(* Logix 5000 project; controller R400_500_XLS vendor 1 type 14 code 216 rev 31.11; software revision 31.01; part 30 of 32 *)
(* tags used below, declared in another part *)
   Alarm : SINT;   // Wait 3 seconds
   CalibData : UDT_SCALE[8];
   Chem_Pump : UDT_CHEM_PUMP[4];   // Chemical Pump flow rate
   FC45_NextMaintDate : DINT[3];   // Next maintenance due date
   FINAL_RINSE_MAX_NBR : INT;   // Maximum nimber of final rinse
   M : DINT[5];   // Memory Bits
   MaxPressRecord : REAL;
   NeutralizantPump : SINT;
   OneShot : DINT[1];
   print_Footer_template : STRING[7];   // Template for the cycle footer
   print_Header_template : STRING[6];   // Template for the cycle header
   PrintCalibdata : STRING[9];
   printNeutralization : STRING[5];
   PrintSensorName : STRING[7];
   printTreatString : STRING[85];   // Treatment String
   rIn_WSH61 : REAL;
   sCRLF : STRING;
   sOut_WSH61 : STRING;
   sPrntArray : STRING[300];   // Printer String Array
   SRE3_Serial_Number : STRING;   // Serial number
   String_Temp : STRING;
   Tmr : TIMER[107];
   WSH41_Total_time : STRING;
   WSH61_Footer : STRING[6];   // The footer being transferred to the print queue.
   CalibCounter : SINT;
   Cfg_11_Modules : BOOL;
   ChemicalName : STRING[9];   // Used by HMI
   CR2Mode : SINT;   // 0= Cycle complete dry contact 1= External pure water valve
   CycleCounter : DINT;
   DateTime : DINT[7];
   ENABLE : BOOL;   // Enable bit
   FC45_NbCycBeforeMaint : DINT;
   iDelayBeforeFillingAuthAlarmMM : DINT;
   iDelayBeforeFillingAuthAlarmSS : DINT;
   iInactivityLogoutTime : DINT;   // Inactivity Logout Time In Minutes
   iPWClosingDelayMM : DINT;
   iPWClosingDelaySS : DINT;
   iSCADACycleCompleteTimeHr : INT;
   iSCADACycleCompleteTimeMin : INT;
   iSCADACycleCompleteTimeSec : INT;
   Language_English : STRING;
   Non_Vented_with_Dry_Option : BOOL;
   NonVented_Without_Dry_Option : BOOL;
   NumInput : UDT_NUMERIC_INPUT[65];   // Numeric input
   NumInputReal : UDT_NUMERIC_INPUT_REAL[17];
   PressureUnit : BOOL;   // Pressure Unit 0=PSIG 1=BAR
   PrintHardware : STRING[29];
   PrintIndex : DINT;
   PrintSystemOption : STRING[29];
   sChangeLanguage : STRING;   // jplv09
   sCycleCounter : STRING;
   SPV_19 : BOOL;   // Screen 80 Enabled/Disabled Pump pressure monitoring
   sTime : STRING;   // String current time
   Tpb : DINT[11];
   Unit : Hrdwre;   // Unit Configuration
   UnLoad : Doors;
   Vented_with_Dry_Option : BOOL;
(* MainProgram, continued *)

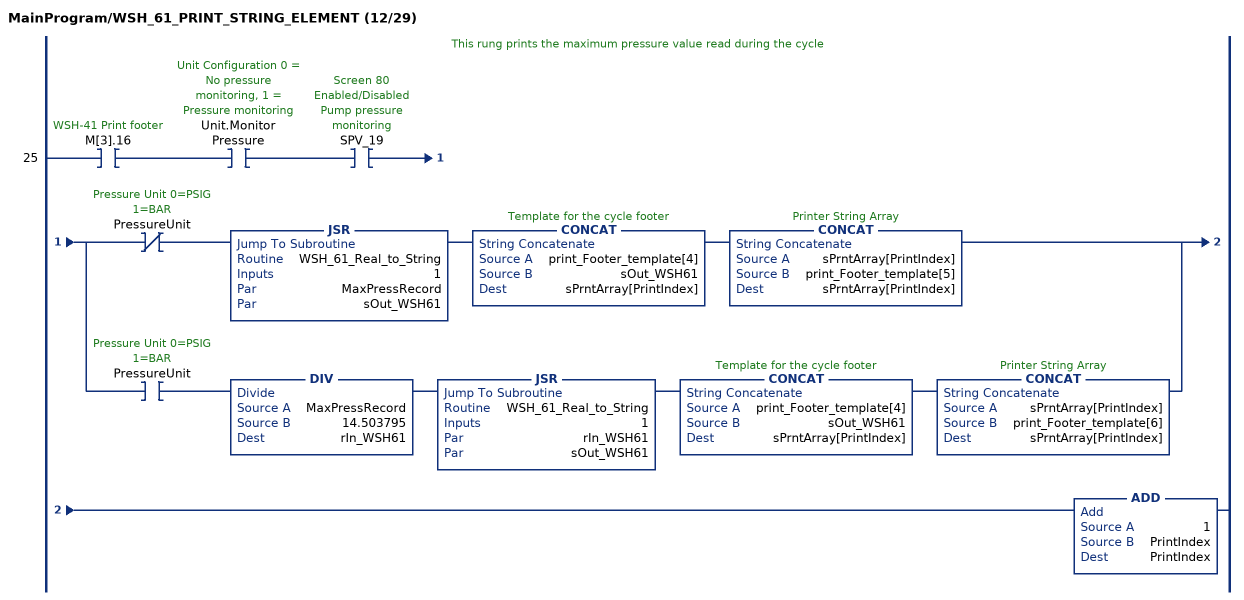
   [picture p617: MainProgram/WSH_61_PRINT_STRING_ELEMENT rungs 25-25]
   // This rung prints the maximum pressure value read during the cycle
   25: XIC(M[3].16)XIC(Unit.MonitorPressure)XIC(SPV_19)[XIO(PressureUnit) JSR(WSH_61_Real_to_String,1,MaxPressRecord,sOut_WSH61) CONCAT(print_Footer_template[4],sOut_WSH61,sPrntArray[PrintIndex]) CONCAT(sPrntArray[PrintIndex],print_Footer_template[5],sPrntArray[PrintIndex]) ,XIC(PressureUnit) DIV(MaxPressRecord,14.503795,rIn_WSH61) JSR(WSH_61_Real_to_String,1,rIn_WSH61,sOut_WSH61) CONCAT(print_Footer_template[4],sOut_WSH61,sPrntArray[PrintIndex]) CONCAT(sPrntArray[PrintIndex],print_Footer_template[6],sPrntArray[PrintIndex]) ]ADD(1,PrintIndex,PrintIndex);
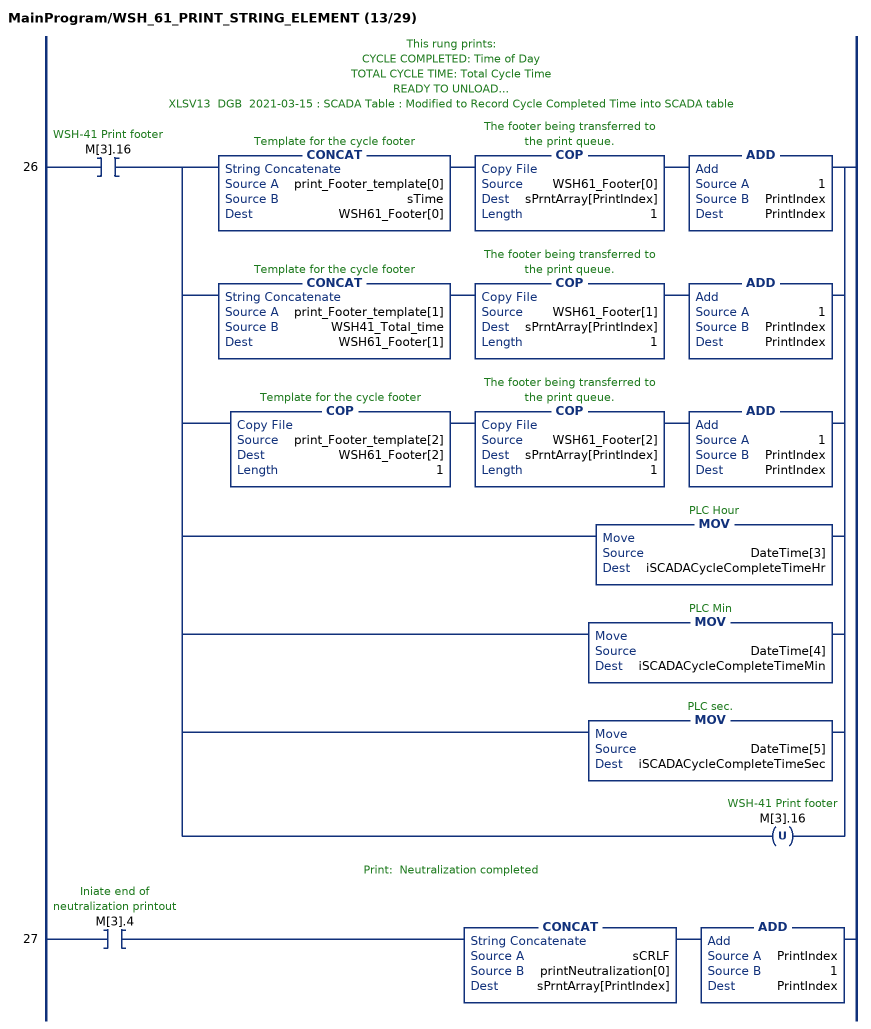
   // This rung prints:
   // CYCLE COMPLETED: Time of Day
   // TOTAL CYCLE TIME: Total Cycle Time
   // READY TO UNLOAD...
   // XLSV13  DGB  2021-03-15 : SCADA Table : Modified to Record Cycle Completed Time into SCADA table
   26: XIC(M[3].16)[CONCAT(print_Footer_template[0],sTime,WSH61_Footer[0]) COP(WSH61_Footer[0],sPrntArray[PrintIndex],1) ADD(1,PrintIndex,PrintIndex) ,CONCAT(print_Footer_template[1],WSH41_Total_time,WSH61_Footer[1]) COP(WSH61_Footer[1],sPrntArray[PrintIndex],1) ADD(1,PrintIndex,PrintIndex) ,COP(print_Footer_template[2],WSH61_Footer[2],1) COP(WSH61_Footer[2],sPrntArray[PrintIndex],1) ADD(1,PrintIndex,PrintIndex) ,[MOV(DateTime[3],iSCADACycleCompleteTimeHr) ,MOV(DateTime[4],iSCADACycleCompleteTimeMin) ,MOV(DateTime[5],iSCADACycleCompleteTimeSec) ] ,OTU(M[3].16) ];
   // Print:  Neutralization completed
   27: XIC(M[3].4)CONCAT(sCRLF,printNeutralization[0],sPrntArray[PrintIndex])ADD(PrintIndex,1,PrintIndex);
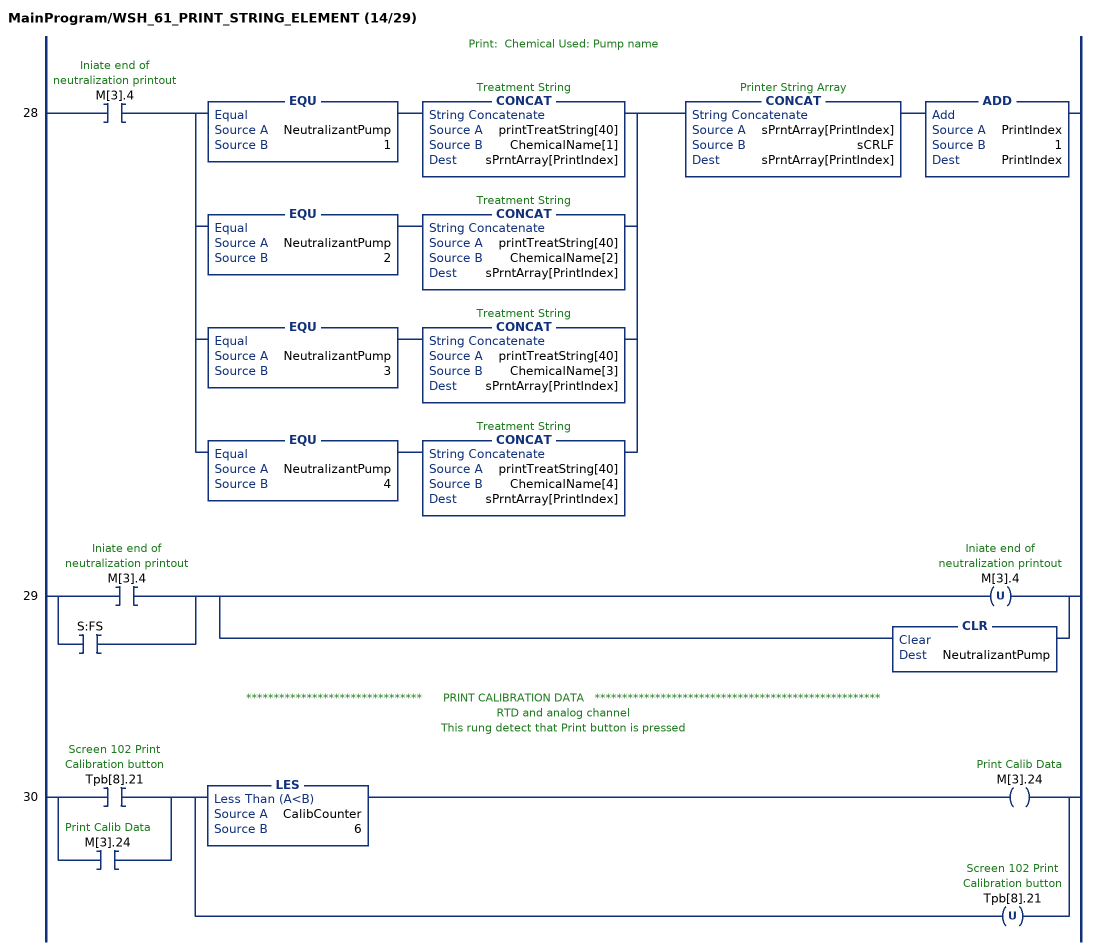
   // Print:  Chemical Used: Pump name
   28: XIC(M[3].4)[EQU(NeutralizantPump,1) CONCAT(printTreatString[40],ChemicalName[1],sPrntArray[PrintIndex]) ,EQU(NeutralizantPump,2) CONCAT(printTreatString[40],ChemicalName[2],sPrntArray[PrintIndex]) ,EQU(NeutralizantPump,3) CONCAT(printTreatString[40],ChemicalName[3],sPrntArray[PrintIndex]) ,EQU(NeutralizantPump,4) CONCAT(printTreatString[40],ChemicalName[4],sPrntArray[PrintIndex]) ]CONCAT(sPrntArray[PrintIndex],sCRLF,sPrntArray[PrintIndex])ADD(PrintIndex,1,PrintIndex);
   29: [XIC(M[3].4) ,XIC(S:FS) ][OTU(M[3].4) ,CLR(NeutralizantPump) ];
   // ********************************      PRINT CALIBRATION DATA   ****************************************************
   // RTD and analog channel
   // This rung detect that Print button is pressed
   30: [XIC(Tpb[8].21) ,XIC(M[3].24) ][LES(CalibCounter,6) OTE(M[3].24) ,OTU(Tpb[8].21) ];
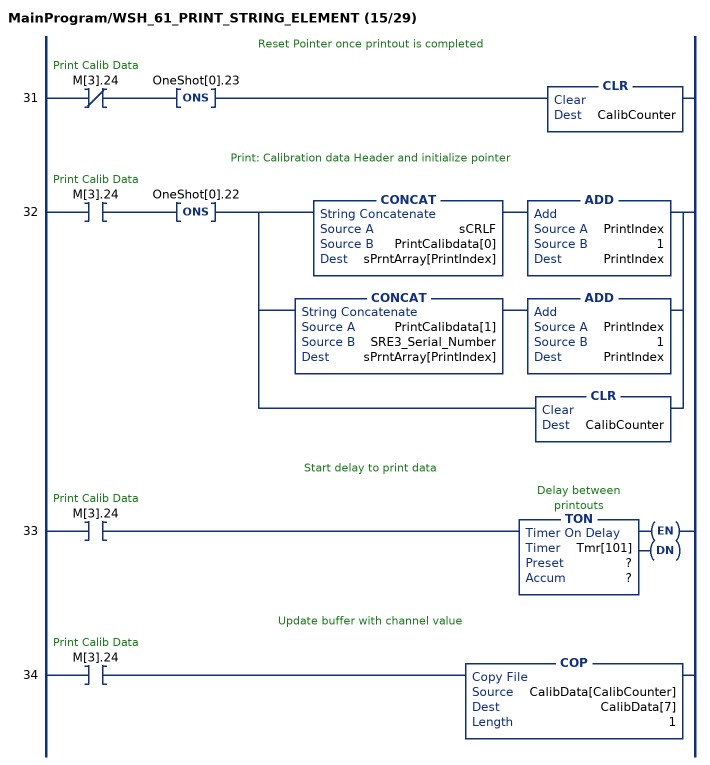
   // Reset Pointer once printout is completed
   31: XIO(M[3].24)ONS(OneShot[0].23)CLR(CalibCounter);
   // Print: Calibration data Header and initialize pointer
   32: XIC(M[3].24)ONS(OneShot[0].22)[CONCAT(sCRLF,PrintCalibdata[0],sPrntArray[PrintIndex]) ADD(PrintIndex,1,PrintIndex) ,CONCAT(PrintCalibdata[1],SRE3_Serial_Number,sPrntArray[PrintIndex]) ADD(PrintIndex,1,PrintIndex) ,CLR(CalibCounter) ];
   // Start delay to print data
   33: XIC(M[3].24)TON(Tmr[101],?,?);
   // Update buffer with channel value
   34: XIC(M[3].24)COP(CalibData[CalibCounter],CalibData[7],1);
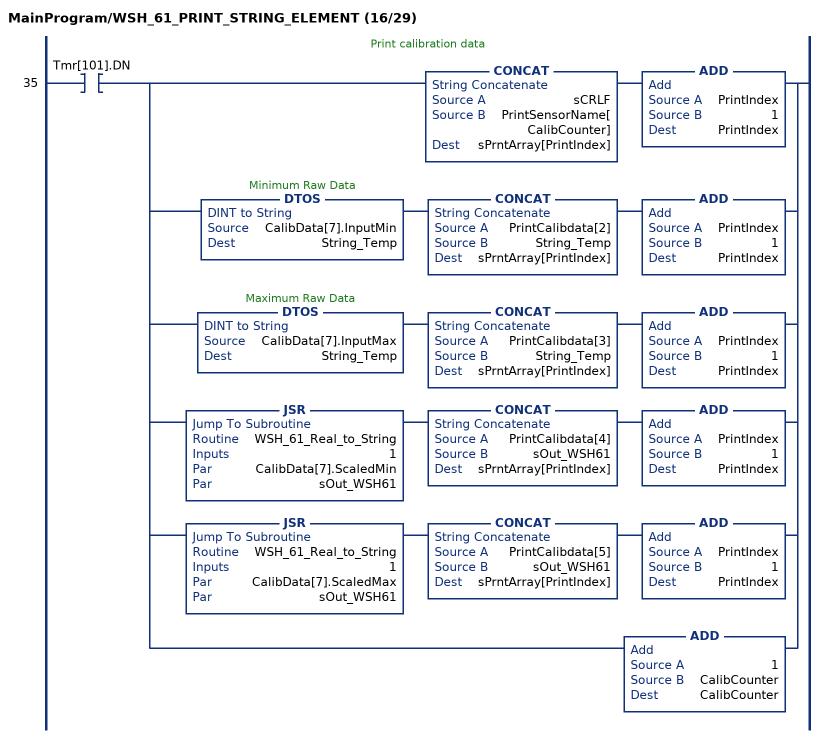
   // Print calibration data
   35: XIC(Tmr[101].DN)[CONCAT(sCRLF,PrintSensorName[CalibCounter],sPrntArray[PrintIndex]) ADD(PrintIndex,1,PrintIndex) ,DTOS(CalibData[7].InputMin,String_Temp) CONCAT(PrintCalibdata[2],String_Temp,sPrntArray[PrintIndex]) ADD(PrintIndex,1,PrintIndex) ,DTOS(CalibData[7].InputMax,String_Temp) CONCAT(PrintCalibdata[3],String_Temp,sPrntArray[PrintIndex]) ADD(PrintIndex,1,PrintIndex) ,JSR(WSH_61_Real_to_String,1,CalibData[7].ScaledMin,sOut_WSH61) CONCAT(PrintCalibdata[4],sOut_WSH61,sPrntArray[PrintIndex]) ADD(PrintIndex,1,PrintIndex) ,JSR(WSH_61_Real_to_String,1,CalibData[7].ScaledMax,sOut_WSH61) CONCAT(PrintCalibdata[5],sOut_WSH61,sPrntArray[PrintIndex]) ADD(PrintIndex,1,PrintIndex) ,ADD(1,CalibCounter,CalibCounter) ];
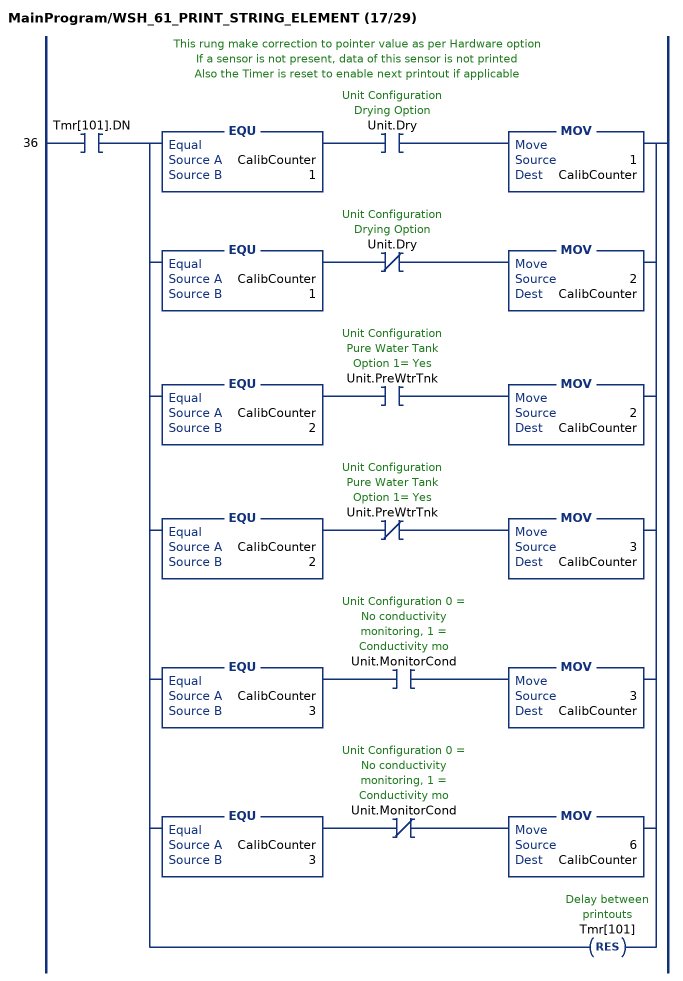
   // This rung make correction to pointer value as per Hardware option
   // If a sensor is not present, data of this sensor is not printed
   // Also the Timer is reset to enable next printout if applicable
   36: XIC(Tmr[101].DN)[EQU(CalibCounter,1) XIC(Unit.Dry) MOV(1,CalibCounter) ,EQU(CalibCounter,1) XIO(Unit.Dry) MOV(2,CalibCounter) ,EQU(CalibCounter,2) XIC(Unit.PreWtrTnk) MOV(2,CalibCounter) ,EQU(CalibCounter,2) XIO(Unit.PreWtrTnk) MOV(3,CalibCounter) ,EQU(CalibCounter,3) XIC(Unit.MonitorCond) MOV(3,CalibCounter) ,EQU(CalibCounter,3) XIO(Unit.MonitorCond) MOV(6,CalibCounter) ,RES(Tmr[101]) ];
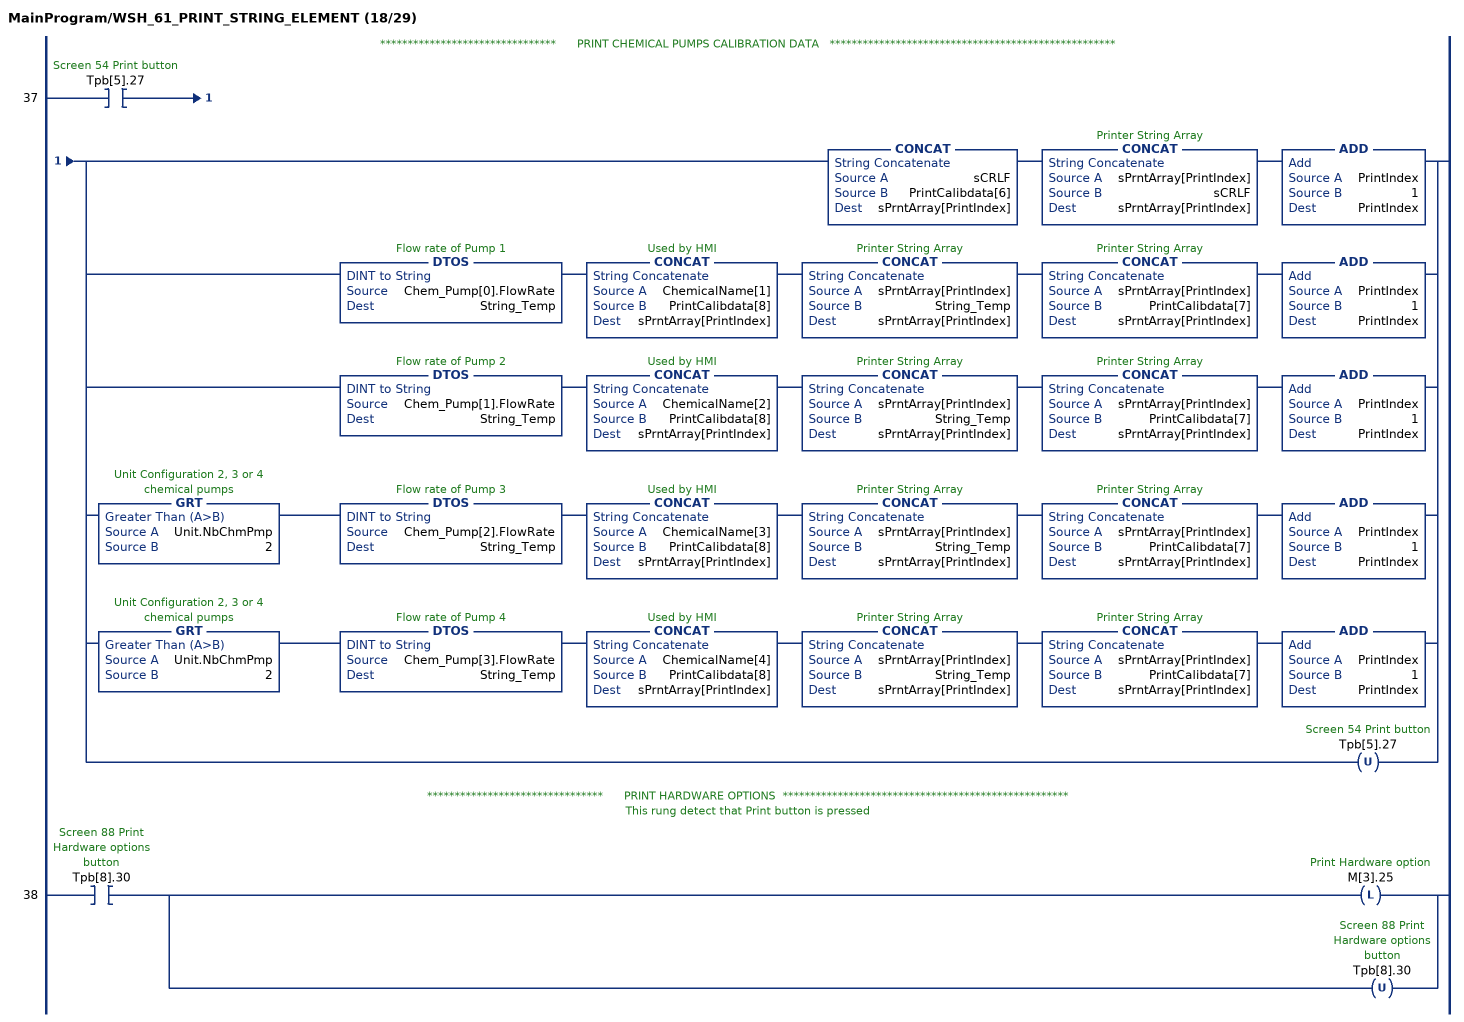
   // ********************************      PRINT CHEMICAL PUMPS CALIBRATION DATA   ****************************************************
   37: XIC(Tpb[5].27)[CONCAT(sCRLF,PrintCalibdata[6],sPrntArray[PrintIndex]) CONCAT(sPrntArray[PrintIndex],sCRLF,sPrntArray[PrintIndex]) ADD(PrintIndex,1,PrintIndex) ,DTOS(Chem_Pump[0].FlowRate,String_Temp) CONCAT(ChemicalName[1],PrintCalibdata[8],sPrntArray[PrintIndex]) CONCAT(sPrntArray[PrintIndex],String_Temp,sPrntArray[PrintIndex]) CONCAT(sPrntArray[PrintIndex],PrintCalibdata[7],sPrntArray[PrintIndex]) ADD(PrintIndex,1,PrintIndex) ,DTOS(Chem_Pump[1].FlowRate,String_Temp) CONCAT(ChemicalName[2],PrintCalibdata[8],sPrntArray[PrintIndex]) CONCAT(sPrntArray[PrintIndex],String_Temp,sPrntArray[PrintIndex]) CONCAT(sPrntArray[PrintIndex],PrintCalibdata[7],sPrntArray[PrintIndex]) ADD(PrintIndex,1,PrintIndex) ,GRT(Unit.NbChmPmp,2) DTOS(Chem_Pump[2].FlowRate,String_Temp) CONCAT(ChemicalName[3],PrintCalibdata[8],sPrntArray[PrintIndex]) CONCAT(sPrntArray[PrintIndex],String_Temp,sPrntArray[PrintIndex]) CONCAT(sPrntArray[PrintIndex],PrintCalibdata[7],sPrntArray[PrintIndex]) ADD(PrintIndex,1,PrintIndex) ,GRT(Unit.NbChmPmp,2) DTOS(Chem_Pump[3].FlowRate,String_Temp) CONCAT(ChemicalName[4],PrintCalibdata[8],sPrntArray[PrintIndex]) CONCAT(sPrntArray[PrintIndex],String_Temp,sPrntArray[PrintIndex]) CONCAT(sPrntArray[PrintIndex],PrintCalibdata[7],sPrntArray[PrintIndex]) ADD(PrintIndex,1,PrintIndex) ,OTU(Tpb[5].27) ];
   // ********************************      PRINT HARDWARE OPTIONS  ****************************************************
   // This rung detect that Print button is pressed
   38: XIC(Tpb[8].30)[OTL(M[3].25) ,OTU(Tpb[8].30) ];
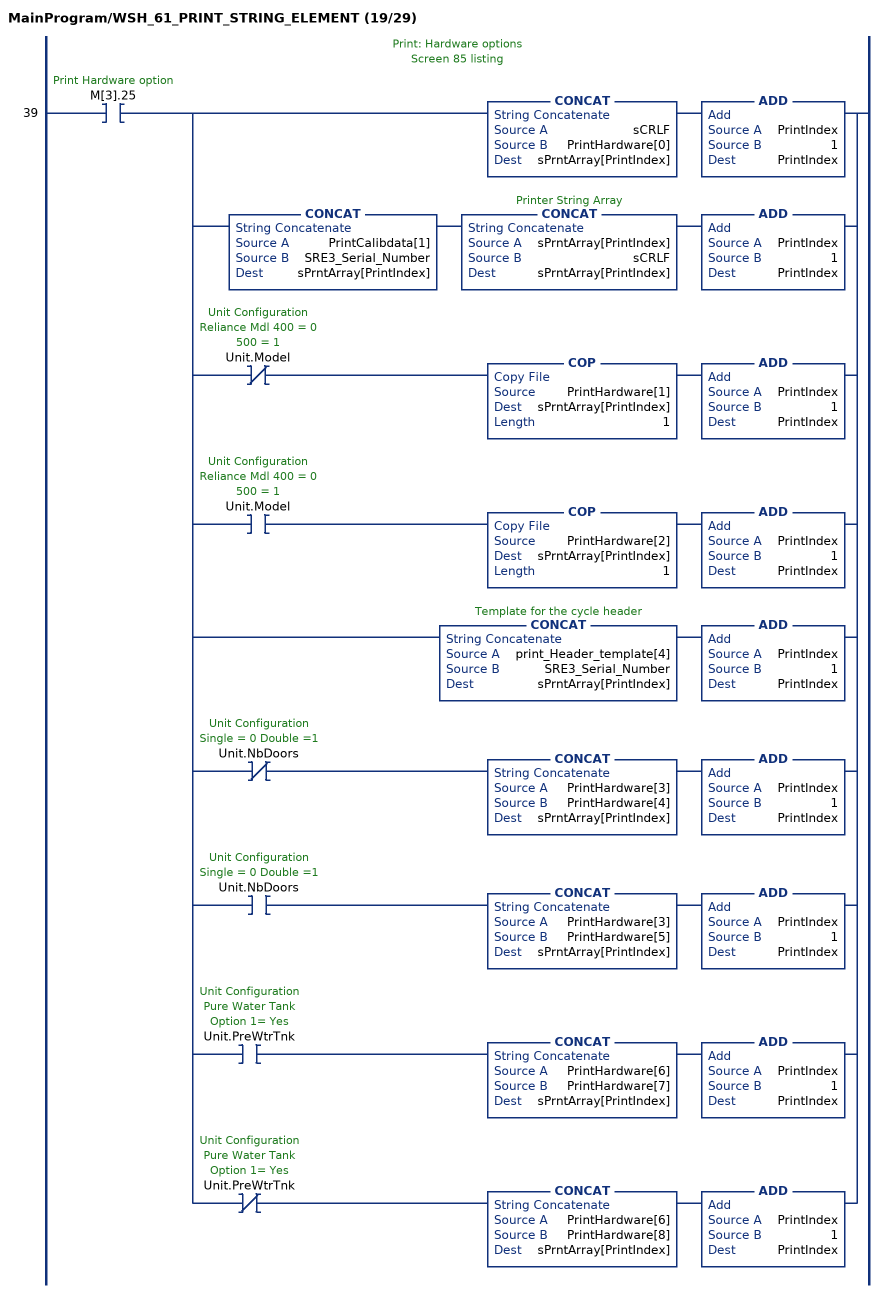
   // Print: Hardware options
   // Screen 85 listing
   39: XIC(M[3].25)[CONCAT(sCRLF,PrintHardware[0],sPrntArray[PrintIndex]) ADD(PrintIndex,1,PrintIndex) ,CONCAT(PrintCalibdata[1],SRE3_Serial_Number,sPrntArray[PrintIndex]) CONCAT(sPrntArray[PrintIndex],sCRLF,sPrntArray[PrintIndex]) ADD(PrintIndex,1,PrintIndex) ,XIO(Unit.Model) COP(PrintHardware[1],sPrntArray[PrintIndex],1) ADD(PrintIndex,1,PrintIndex) ,XIC(Unit.Model) COP(PrintHardware[2],sPrntArray[PrintIndex],1) ADD(PrintIndex,1,PrintIndex) ,CONCAT(print_Header_template[4],SRE3_Serial_Number,sPrntArray[PrintIndex]) ADD(PrintIndex,1,PrintIndex) ,XIO(Unit.NbDoors) CONCAT(PrintHardware[3],PrintHardware[4],sPrntArray[PrintIndex]) ADD(PrintIndex,1,PrintIndex) ,XIC(Unit.NbDoors) CONCAT(PrintHardware[3],PrintHardware[5],sPrntArray[PrintIndex]) ADD(PrintIndex,1,PrintIndex) ,XIC(Unit.PreWtrTnk) CONCAT(PrintHardware[6],PrintHardware[7],sPrntArray[PrintIndex]) ADD(PrintIndex,1,PrintIndex) ,XIO(Unit.PreWtrTnk) CONCAT(PrintHardware[6],PrintHardware[8],sPrntArray[PrintIndex]) ADD(PrintIndex,1,PrintIndex) ];
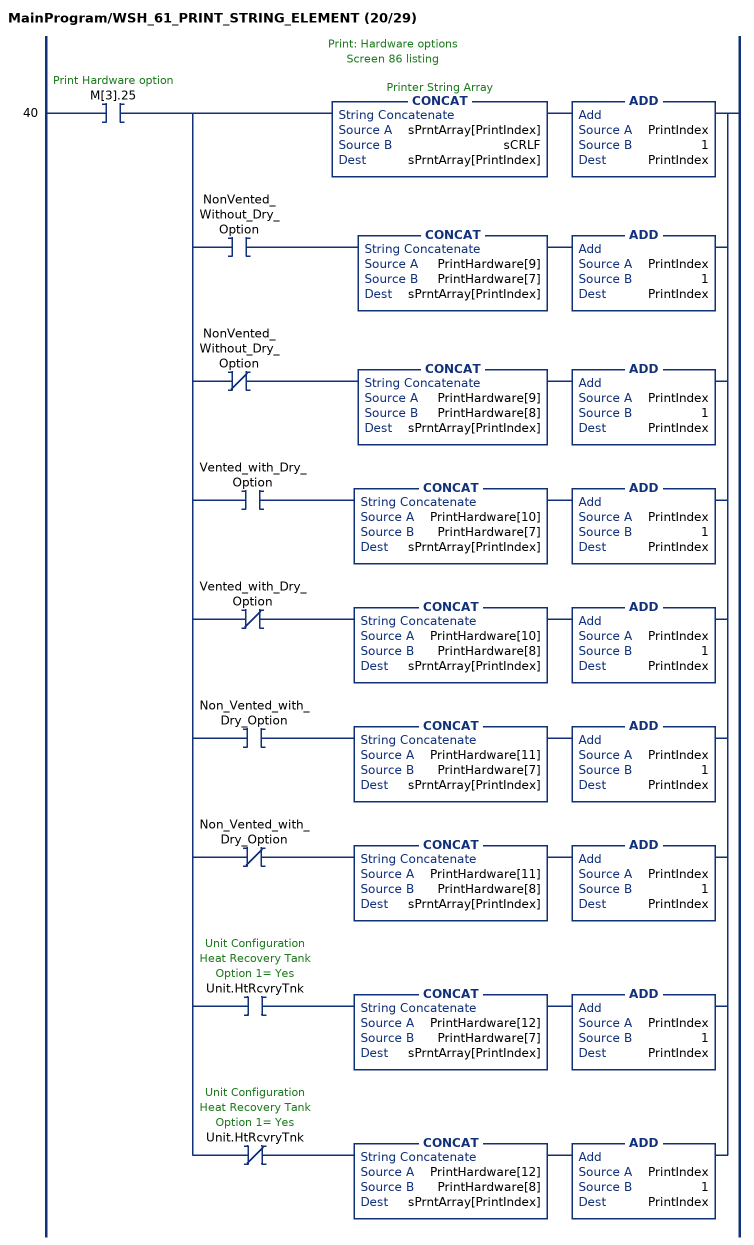
   // Print: Hardware options
   // Screen 86 listing
   40: XIC(M[3].25)[CONCAT(sPrntArray[PrintIndex],sCRLF,sPrntArray[PrintIndex]) ADD(PrintIndex,1,PrintIndex) ,XIC(NonVented_Without_Dry_Option) CONCAT(PrintHardware[9],PrintHardware[7],sPrntArray[PrintIndex]) ADD(PrintIndex,1,PrintIndex) ,XIO(NonVented_Without_Dry_Option) CONCAT(PrintHardware[9],PrintHardware[8],sPrntArray[PrintIndex]) ADD(PrintIndex,1,PrintIndex) ,XIC(Vented_with_Dry_Option) CONCAT(PrintHardware[10],PrintHardware[7],sPrntArray[PrintIndex]) ADD(PrintIndex,1,PrintIndex) ,XIO(Vented_with_Dry_Option) CONCAT(PrintHardware[10],PrintHardware[8],sPrntArray[PrintIndex]) ADD(PrintIndex,1,PrintIndex) ,XIC(Non_Vented_with_Dry_Option) CONCAT(PrintHardware[11],PrintHardware[7],sPrntArray[PrintIndex]) ADD(PrintIndex,1,PrintIndex) ,XIO(Non_Vented_with_Dry_Option) CONCAT(PrintHardware[11],PrintHardware[8],sPrntArray[PrintIndex]) ADD(PrintIndex,1,PrintIndex) ,XIC(Unit.HtRcvryTnk) CONCAT(PrintHardware[12],PrintHardware[7],sPrntArray[PrintIndex]) ADD(PrintIndex,1,PrintIndex) ,XIO(Unit.HtRcvryTnk) CONCAT(PrintHardware[12],PrintHardware[8],sPrntArray[PrintIndex]) ADD(PrintIndex,1,PrintIndex) ];
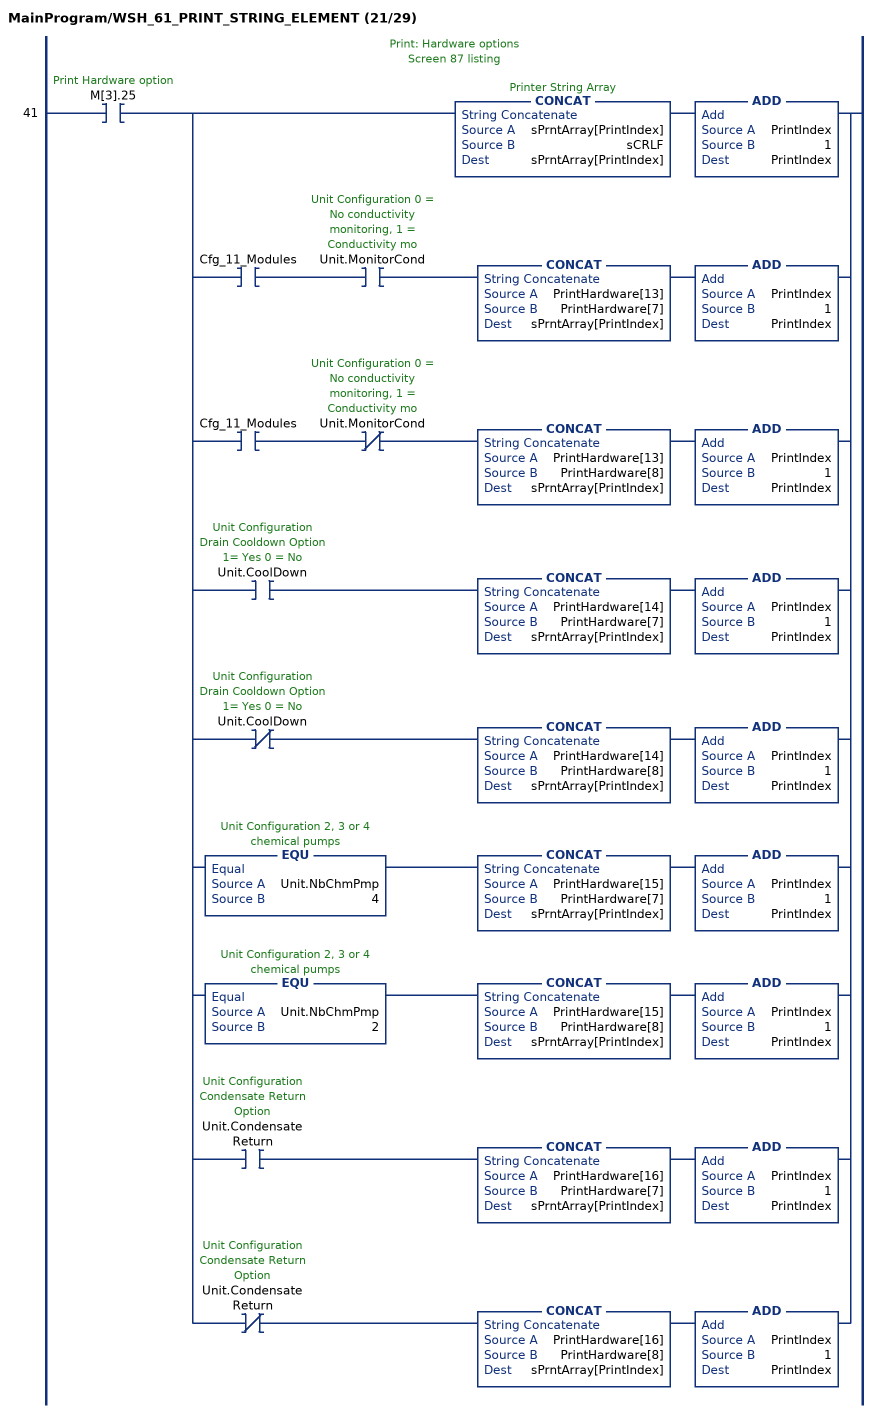
   // Print: Hardware options
   // Screen 87 listing
   41: XIC(M[3].25)[CONCAT(sPrntArray[PrintIndex],sCRLF,sPrntArray[PrintIndex]) ADD(PrintIndex,1,PrintIndex) ,XIC(Cfg_11_Modules) XIC(Unit.MonitorCond) CONCAT(PrintHardware[13],PrintHardware[7],sPrntArray[PrintIndex]) ADD(PrintIndex,1,PrintIndex) ,XIC(Cfg_11_Modules) XIO(Unit.MonitorCond) CONCAT(PrintHardware[13],PrintHardware[8],sPrntArray[PrintIndex]) ADD(PrintIndex,1,PrintIndex) ,XIC(Unit.CoolDown) CONCAT(PrintHardware[14],PrintHardware[7],sPrntArray[PrintIndex]) ADD(PrintIndex,1,PrintIndex) ,XIO(Unit.CoolDown) CONCAT(PrintHardware[14],PrintHardware[8],sPrntArray[PrintIndex]) ADD(PrintIndex,1,PrintIndex) ,EQU(Unit.NbChmPmp,4) CONCAT(PrintHardware[15],PrintHardware[7],sPrntArray[PrintIndex]) ADD(PrintIndex,1,PrintIndex) ,EQU(Unit.NbChmPmp,2) CONCAT(PrintHardware[15],PrintHardware[8],sPrntArray[PrintIndex]) ADD(PrintIndex,1,PrintIndex) ,XIC(Unit.CondensateReturn) CONCAT(PrintHardware[16],PrintHardware[7],sPrntArray[PrintIndex]) ADD(PrintIndex,1,PrintIndex) ,XIO(Unit.CondensateReturn) CONCAT(PrintHardware[16],PrintHardware[8],sPrntArray[PrintIndex]) ADD(PrintIndex,1,PrintIndex) ];
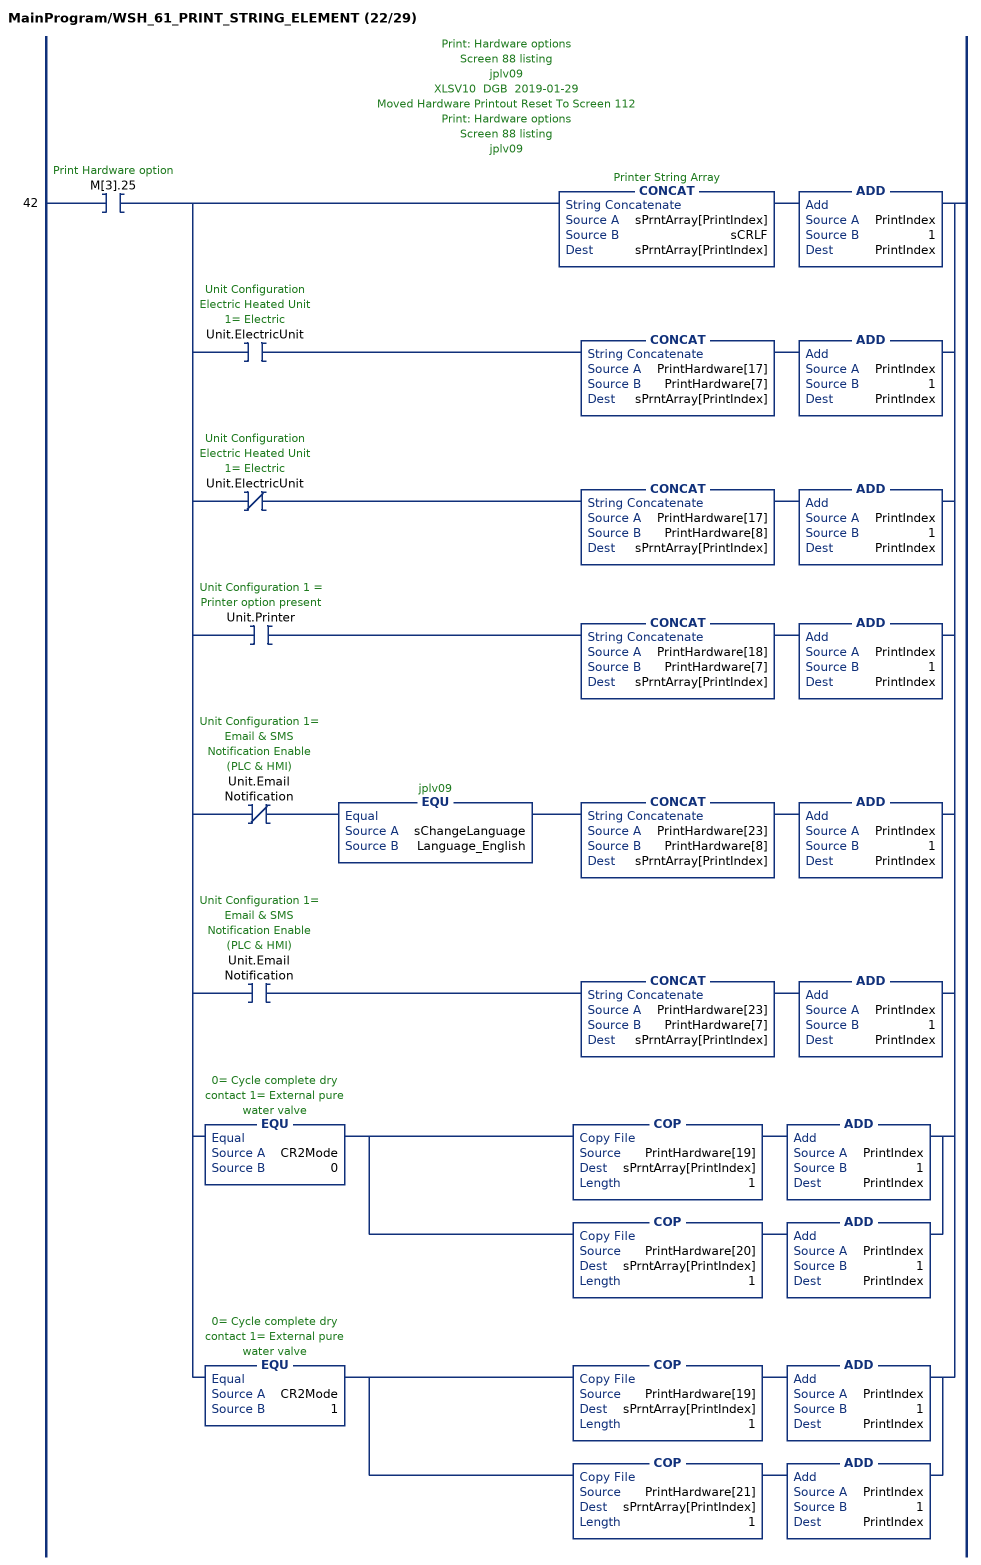
   // Print: Hardware options
   // Screen 88 listing
   // jplv09
   // XLSV10  DGB  2019-01-29
   // Moved Hardware Printout Reset To Screen 112
   // Print: Hardware options
   // Screen 88 listing
   // jplv09
   42: XIC(M[3].25)[CONCAT(sPrntArray[PrintIndex],sCRLF,sPrntArray[PrintIndex]) ADD(PrintIndex,1,PrintIndex) ,XIC(Unit.ElectricUnit) CONCAT(PrintHardware[17],PrintHardware[7],sPrntArray[PrintIndex]) ADD(PrintIndex,1,PrintIndex) ,XIO(Unit.ElectricUnit) CONCAT(PrintHardware[17],PrintHardware[8],sPrntArray[PrintIndex]) ADD(PrintIndex,1,PrintIndex) ,XIC(Unit.Printer) CONCAT(PrintHardware[18],PrintHardware[7],sPrntArray[PrintIndex]) ADD(PrintIndex,1,PrintIndex) ,XIO(Unit.EmailNotification) EQU(sChangeLanguage,Language_English) CONCAT(PrintHardware[23],PrintHardware[8],sPrntArray[PrintIndex]) ADD(PrintIndex,1,PrintIndex) ,XIC(Unit.EmailNotification) CONCAT(PrintHardware[23],PrintHardware[7],sPrntArray[PrintIndex]) ADD(PrintIndex,1,PrintIndex) ,EQU(CR2Mode,0) [COP(PrintHardware[19],sPrntArray[PrintIndex],1) ADD(PrintIndex,1,PrintIndex) ,COP(PrintHardware[20],sPrntArray[PrintIndex],1) ADD(PrintIndex,1,PrintIndex) ] ,EQU(CR2Mode,1) [COP(PrintHardware[19],sPrntArray[PrintIndex],1) ADD(PrintIndex,1,PrintIndex) ,COP(PrintHardware[21],sPrntArray[PrintIndex],1) ADD(PrintIndex,1,PrintIndex) ] ];
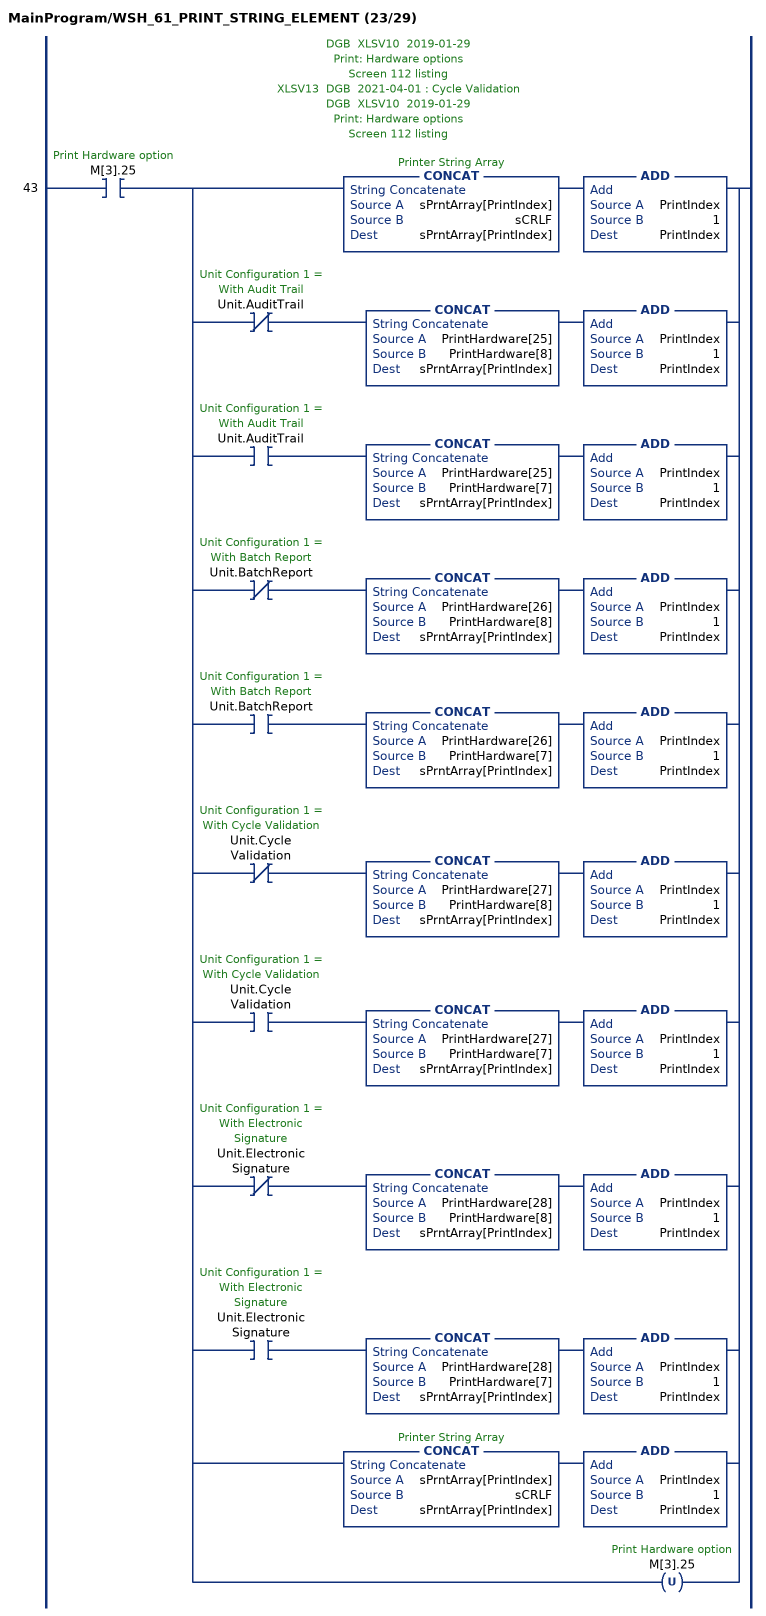
   // DGB  XLSV10  2019-01-29
   // Print: Hardware options
   // Screen 112 listing
   // XLSV13  DGB  2021-04-01 : Cycle Validation
   // DGB  XLSV10  2019-01-29
   // Print: Hardware options
   // Screen 112 listing
   43: XIC(M[3].25)[CONCAT(sPrntArray[PrintIndex],sCRLF,sPrntArray[PrintIndex]) ADD(PrintIndex,1,PrintIndex) ,XIO(Unit.AuditTrail) CONCAT(PrintHardware[25],PrintHardware[8],sPrntArray[PrintIndex]) ADD(PrintIndex,1,PrintIndex) ,XIC(Unit.AuditTrail) CONCAT(PrintHardware[25],PrintHardware[7],sPrntArray[PrintIndex]) ADD(PrintIndex,1,PrintIndex) ,XIO(Unit.BatchReport) CONCAT(PrintHardware[26],PrintHardware[8],sPrntArray[PrintIndex]) ADD(PrintIndex,1,PrintIndex) ,XIC(Unit.BatchReport) CONCAT(PrintHardware[26],PrintHardware[7],sPrntArray[PrintIndex]) ADD(PrintIndex,1,PrintIndex) ,XIO(Unit.CycleValidation) CONCAT(PrintHardware[27],PrintHardware[8],sPrntArray[PrintIndex]) ADD(PrintIndex,1,PrintIndex) ,XIC(Unit.CycleValidation) CONCAT(PrintHardware[27],PrintHardware[7],sPrntArray[PrintIndex]) ADD(PrintIndex,1,PrintIndex) ,XIO(Unit.ElectronicSignature) CONCAT(PrintHardware[28],PrintHardware[8],sPrntArray[PrintIndex]) ADD(PrintIndex,1,PrintIndex) ,XIC(Unit.ElectronicSignature) CONCAT(PrintHardware[28],PrintHardware[7],sPrntArray[PrintIndex]) ADD(PrintIndex,1,PrintIndex) ,CONCAT(sPrntArray[PrintIndex],sCRLF,sPrntArray[PrintIndex]) ADD(PrintIndex,1,PrintIndex) ,OTU(M[3].25) ];
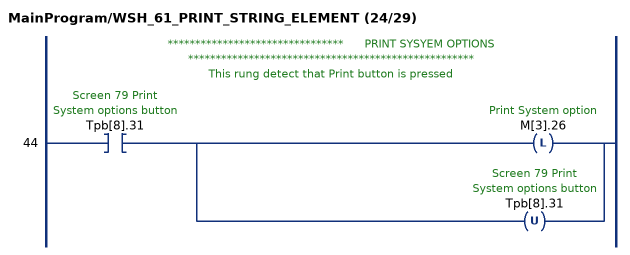
   // ********************************      PRINT SYSYEM OPTIONS  ****************************************************
   // This rung detect that Print button is pressed
   44: XIC(Tpb[8].31)[OTL(M[3].26) ,OTU(Tpb[8].31) ];
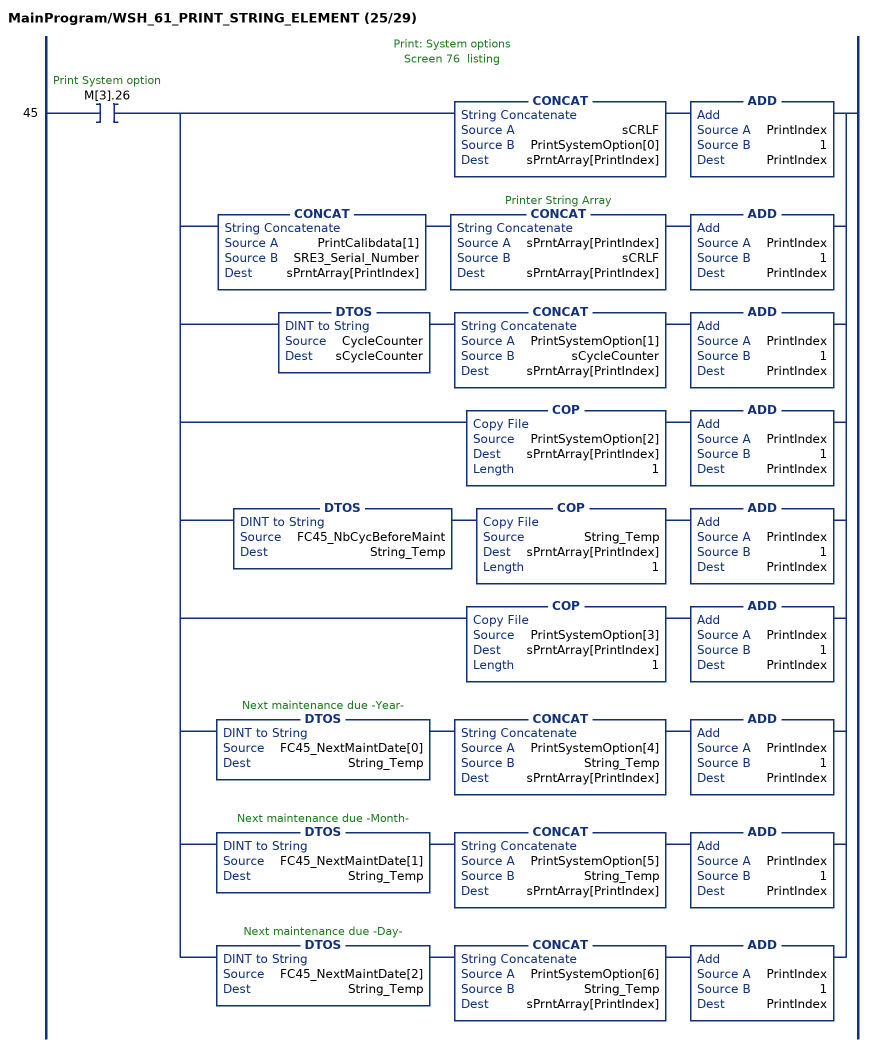
   // Print: System options
   // Screen 76  listing
   45: XIC(M[3].26)[CONCAT(sCRLF,PrintSystemOption[0],sPrntArray[PrintIndex]) ADD(PrintIndex,1,PrintIndex) ,CONCAT(PrintCalibdata[1],SRE3_Serial_Number,sPrntArray[PrintIndex]) CONCAT(sPrntArray[PrintIndex],sCRLF,sPrntArray[PrintIndex]) ADD(PrintIndex,1,PrintIndex) ,DTOS(CycleCounter,sCycleCounter) CONCAT(PrintSystemOption[1],sCycleCounter,sPrntArray[PrintIndex]) ADD(PrintIndex,1,PrintIndex) ,COP(PrintSystemOption[2],sPrntArray[PrintIndex],1) ADD(PrintIndex,1,PrintIndex) ,DTOS(FC45_NbCycBeforeMaint,String_Temp) COP(String_Temp,sPrntArray[PrintIndex],1) ADD(PrintIndex,1,PrintIndex) ,COP(PrintSystemOption[3],sPrntArray[PrintIndex],1) ADD(PrintIndex,1,PrintIndex) ,DTOS(FC45_NextMaintDate[0],String_Temp) CONCAT(PrintSystemOption[4],String_Temp,sPrntArray[PrintIndex]) ADD(PrintIndex,1,PrintIndex) ,DTOS(FC45_NextMaintDate[1],String_Temp) CONCAT(PrintSystemOption[5],String_Temp,sPrntArray[PrintIndex]) ADD(PrintIndex,1,PrintIndex) ,DTOS(FC45_NextMaintDate[2],String_Temp) CONCAT(PrintSystemOption[6],String_Temp,sPrntArray[PrintIndex]) ADD(PrintIndex,1,PrintIndex) ];
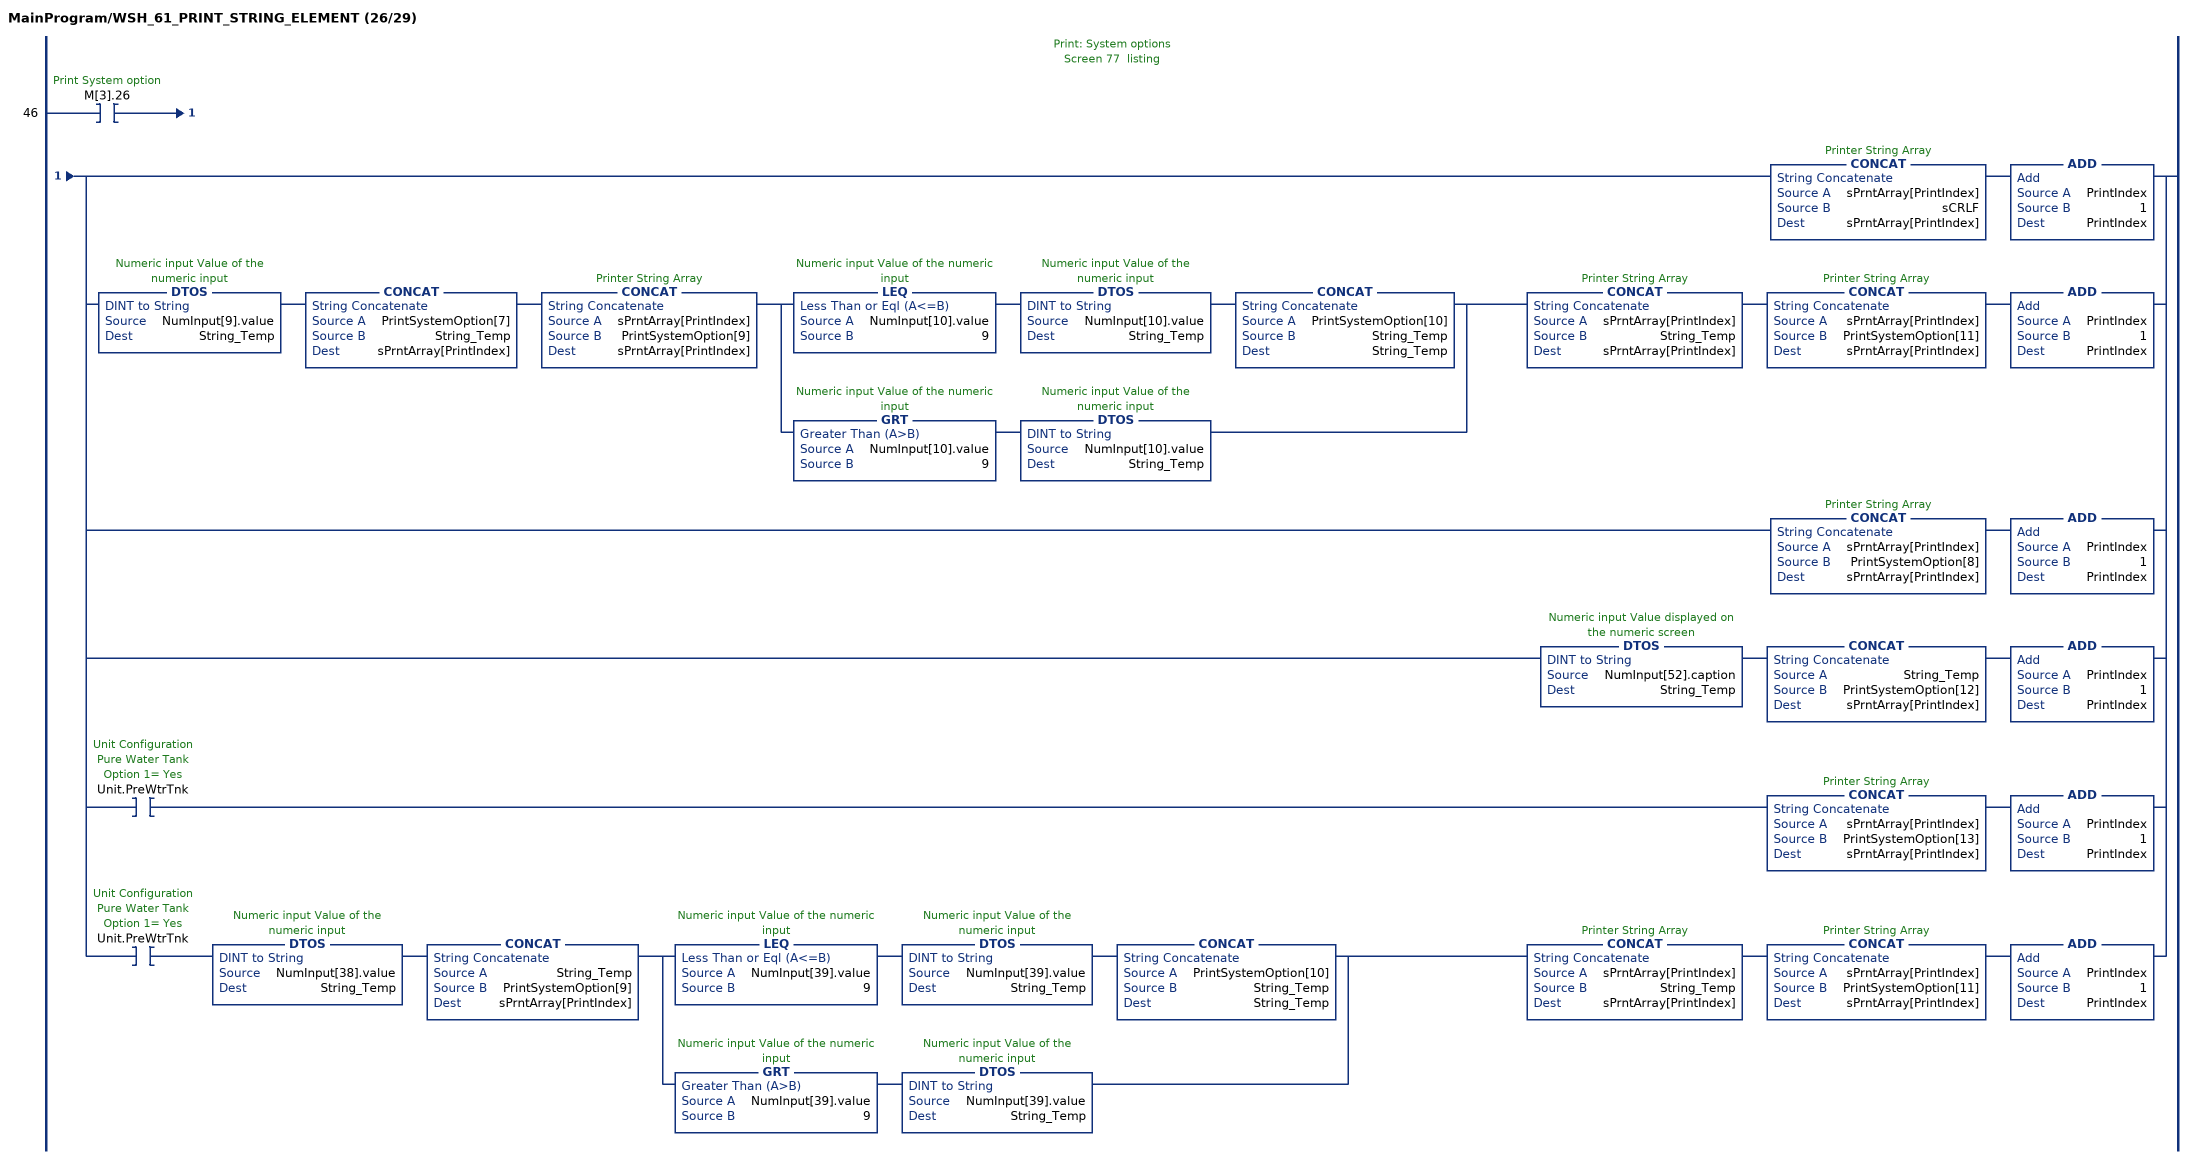
   // Print: System options
   // Screen 77  listing
   46: XIC(M[3].26)[CONCAT(sPrntArray[PrintIndex],sCRLF,sPrntArray[PrintIndex]) ADD(PrintIndex,1,PrintIndex) ,DTOS(NumInput[9].value,String_Temp) CONCAT(PrintSystemOption[7],String_Temp,sPrntArray[PrintIndex]) CONCAT(sPrntArray[PrintIndex],PrintSystemOption[9],sPrntArray[PrintIndex]) [LEQ(NumInput[10].value,9) DTOS(NumInput[10].value,String_Temp) CONCAT(PrintSystemOption[10],String_Temp,String_Temp) ,GRT(NumInput[10].value,9) DTOS(NumInput[10].value,String_Temp) ] CONCAT(sPrntArray[PrintIndex],String_Temp,sPrntArray[PrintIndex]) CONCAT(sPrntArray[PrintIndex],PrintSystemOption[11],sPrntArray[PrintIndex]) ADD(PrintIndex,1,PrintIndex) ,CONCAT(sPrntArray[PrintIndex],PrintSystemOption[8],sPrntArray[PrintIndex]) ADD(PrintIndex,1,PrintIndex) ,DTOS(NumInput[52].caption,String_Temp) CONCAT(String_Temp,PrintSystemOption[12],sPrntArray[PrintIndex]) ADD(PrintIndex,1,PrintIndex) ,XIC(Unit.PreWtrTnk) CONCAT(sPrntArray[PrintIndex],PrintSystemOption[13],sPrntArray[PrintIndex]) ADD(PrintIndex,1,PrintIndex) ,XIC(Unit.PreWtrTnk) DTOS(NumInput[38].value,String_Temp) CONCAT(String_Temp,PrintSystemOption[9],sPrntArray[PrintIndex]) [LEQ(NumInput[39].value,9) DTOS(NumInput[39].value,String_Temp) CONCAT(PrintSystemOption[10],String_Temp,String_Temp) ,GRT(NumInput[39].value,9) DTOS(NumInput[39].value,String_Temp) ] CONCAT(sPrntArray[PrintIndex],String_Temp,sPrntArray[PrintIndex]) CONCAT(sPrntArray[PrintIndex],PrintSystemOption[11],sPrntArray[PrintIndex]) ADD(PrintIndex,1,PrintIndex) ];
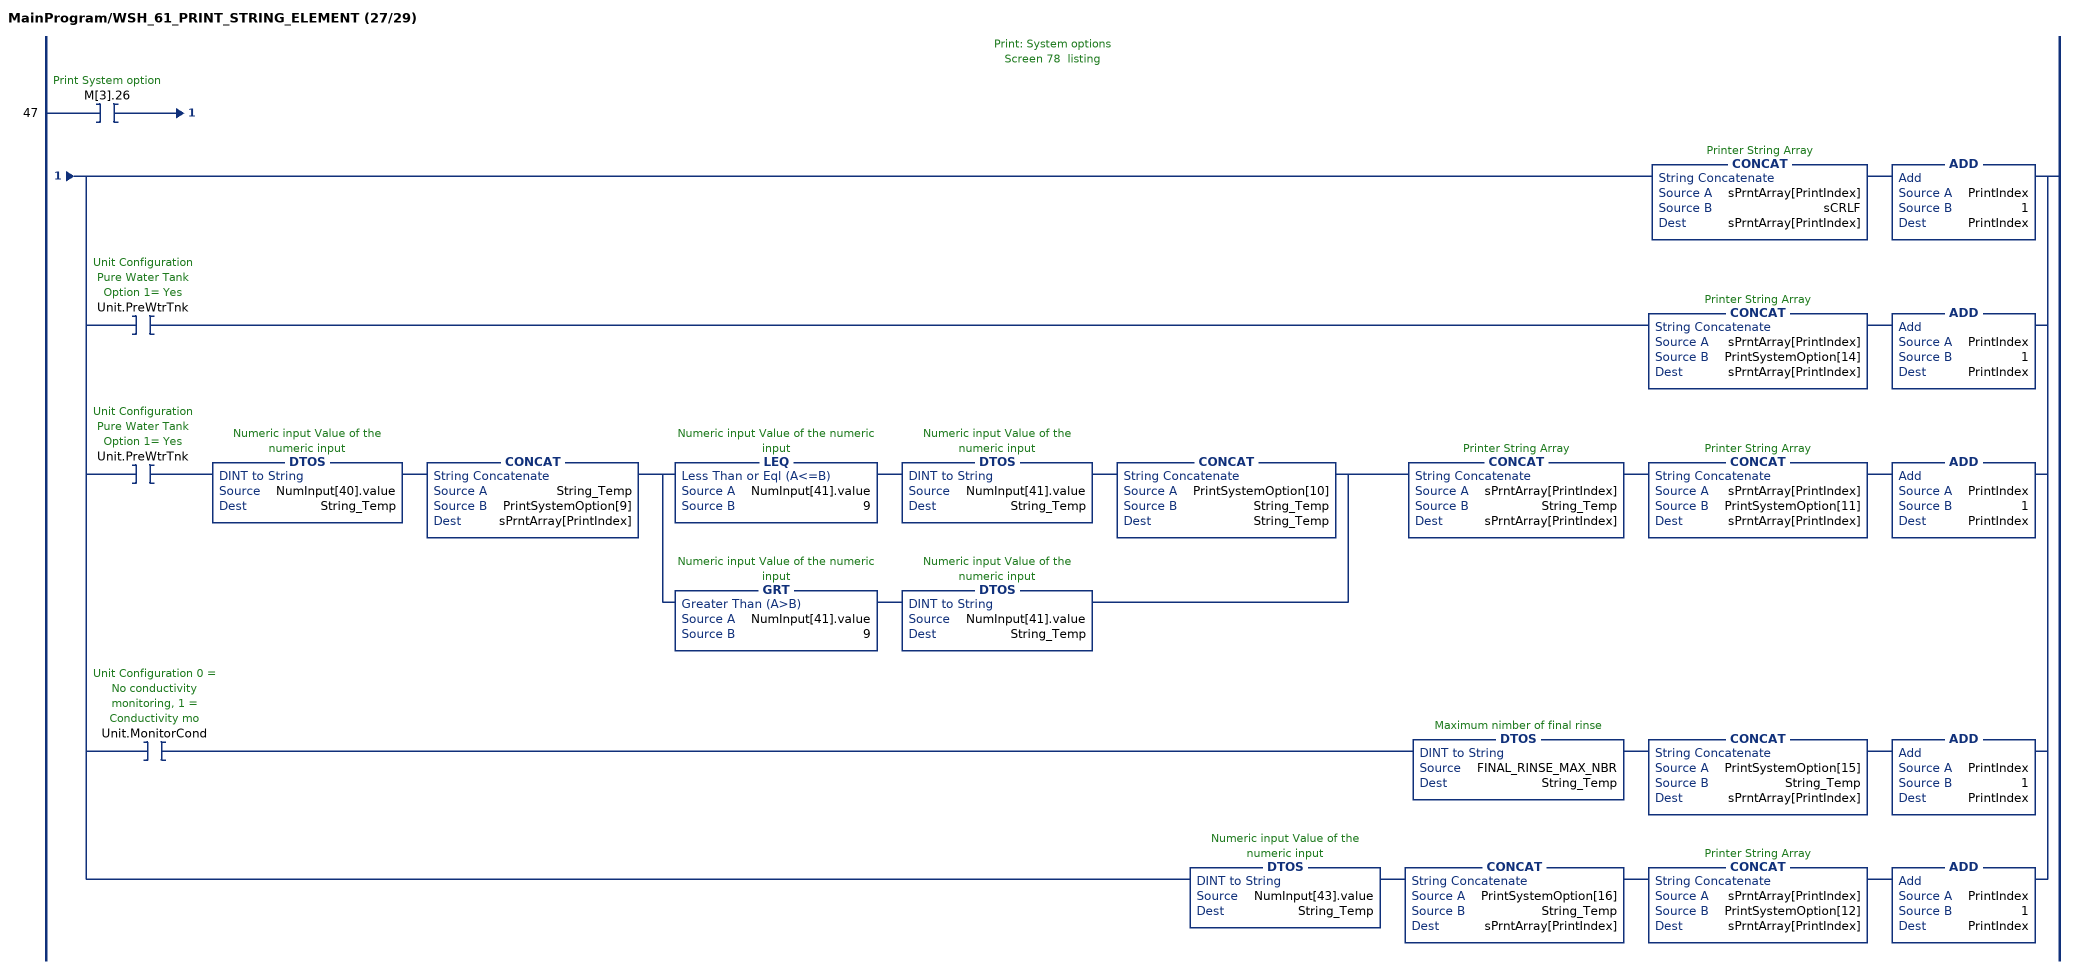
   // Print: System options
   // Screen 78  listing
   47: XIC(M[3].26)[CONCAT(sPrntArray[PrintIndex],sCRLF,sPrntArray[PrintIndex]) ADD(PrintIndex,1,PrintIndex) ,XIC(Unit.PreWtrTnk) CONCAT(sPrntArray[PrintIndex],PrintSystemOption[14],sPrntArray[PrintIndex]) ADD(PrintIndex,1,PrintIndex) ,XIC(Unit.PreWtrTnk) DTOS(NumInput[40].value,String_Temp) CONCAT(String_Temp,PrintSystemOption[9],sPrntArray[PrintIndex]) [LEQ(NumInput[41].value,9) DTOS(NumInput[41].value,String_Temp) CONCAT(PrintSystemOption[10],String_Temp,String_Temp) ,GRT(NumInput[41].value,9) DTOS(NumInput[41].value,String_Temp) ] CONCAT(sPrntArray[PrintIndex],String_Temp,sPrntArray[PrintIndex]) CONCAT(sPrntArray[PrintIndex],PrintSystemOption[11],sPrntArray[PrintIndex]) ADD(PrintIndex,1,PrintIndex) ,XIC(Unit.MonitorCond) DTOS(FINAL_RINSE_MAX_NBR,String_Temp) CONCAT(PrintSystemOption[15],String_Temp,sPrntArray[PrintIndex]) ADD(PrintIndex,1,PrintIndex) ,DTOS(NumInput[43].value,String_Temp) CONCAT(PrintSystemOption[16],String_Temp,sPrntArray[PrintIndex]) CONCAT(sPrntArray[PrintIndex],PrintSystemOption[12],sPrntArray[PrintIndex]) ADD(PrintIndex,1,PrintIndex) ];
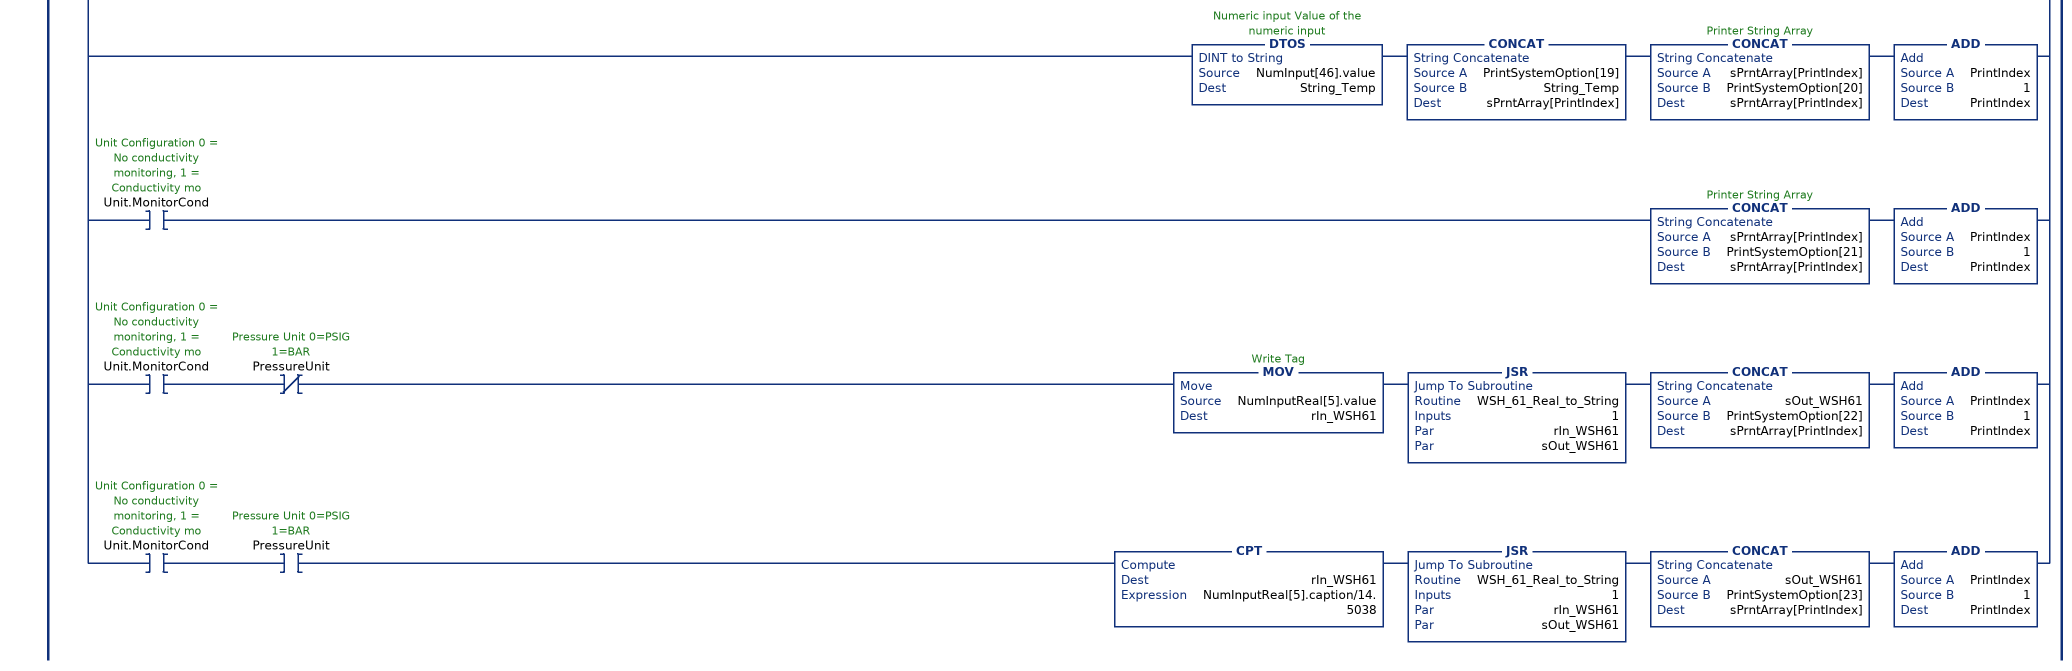
   // Print: System options
   // Screen 79  listing
   // XLSV10  DGB  2019-01-29
   // Moved End of System Option Printout in Screen 114
   48: XIC(M[3].26)[CONCAT(sPrntArray[PrintIndex],sCRLF,sPrntArray[PrintIndex]) ADD(PrintIndex,1,PrintIndex) ,CONCAT(sPrntArray[PrintIndex],PrintSystemOption[17],sPrntArray[PrintIndex]) ADD(PrintIndex,1,PrintIndex) ,DTOS(NumInput[44].value,String_Temp) CONCAT(String_Temp,PrintSystemOption[9],sPrntArray[PrintIndex]) [LEQ(NumInput[45].value,9) DTOS(NumInput[45].value,String_Temp) CONCAT(PrintSystemOption[10],String_Temp,String_Temp) ,GRT(NumInput[45].value,9) DTOS(NumInput[45].value,String_Temp) ] CONCAT(sPrntArray[PrintIndex],String_Temp,sPrntArray[PrintIndex]) CONCAT(sPrntArray[PrintIndex],PrintSystemOption[11],sPrntArray[PrintIndex]) ADD(PrintIndex,1,PrintIndex) ,XIC(Unit.Dry) CONCAT(sPrntArray[PrintIndex],PrintSystemOption[18],sPrntArray[PrintIndex]) ADD(PrintIndex,1,PrintIndex) ,XIC(Unit.Dry) DTOS(NumInput[47].value,String_Temp) CONCAT(String_Temp,PrintSystemOption[9],sPrntArray[PrintIndex]) [LEQ(NumInput[48].value,9) DTOS(NumInput[48].value,String_Temp) CONCAT(PrintSystemOption[10],String_Temp,String_Temp) ,GRT(NumInput[48].value,9) DTOS(NumInput[48].value,String_Temp) ] CONCAT(sPrntArray[PrintIndex],String_Temp,sPrntArray[PrintIndex]) CONCAT(sPrntArray[PrintIndex],PrintSystemOption[11],sPrntArray[PrintIndex]) ADD(PrintIndex,1,PrintIndex) ,DTOS(NumInput[46].value,String_Temp) CONCAT(PrintSystemOption[19],String_Temp,sPrntArray[PrintIndex]) CONCAT(sPrntArray[PrintIndex],PrintSystemOption[20],sPrntArray[PrintIndex]) ADD(PrintIndex,1,PrintIndex) ,XIC(Unit.MonitorCond) CONCAT(sPrntArray[PrintIndex],PrintSystemOption[21],sPrntArray[PrintIndex]) ADD(PrintIndex,1,PrintIndex) ,XIC(Unit.MonitorCond) XIO(PressureUnit) MOV(NumInputReal[5].value,rIn_WSH61) JSR(WSH_61_Real_to_String,1,rIn_WSH61,sOut_WSH61) CONCAT(sOut_WSH61,PrintSystemOption[22],sPrntArray[PrintIndex]) ADD(PrintIndex,1,PrintIndex) ,XIC(Unit.MonitorCond) XIC(PressureUnit) CPT(rIn_WSH61,NumInputReal[5].caption/14.5038) JSR(WSH_61_Real_to_String,1,rIn_WSH61,sOut_WSH61) CONCAT(sOut_WSH61,PrintSystemOption[23],sPrntArray[PrintIndex]) ADD(PrintIndex,1,PrintIndex) ];
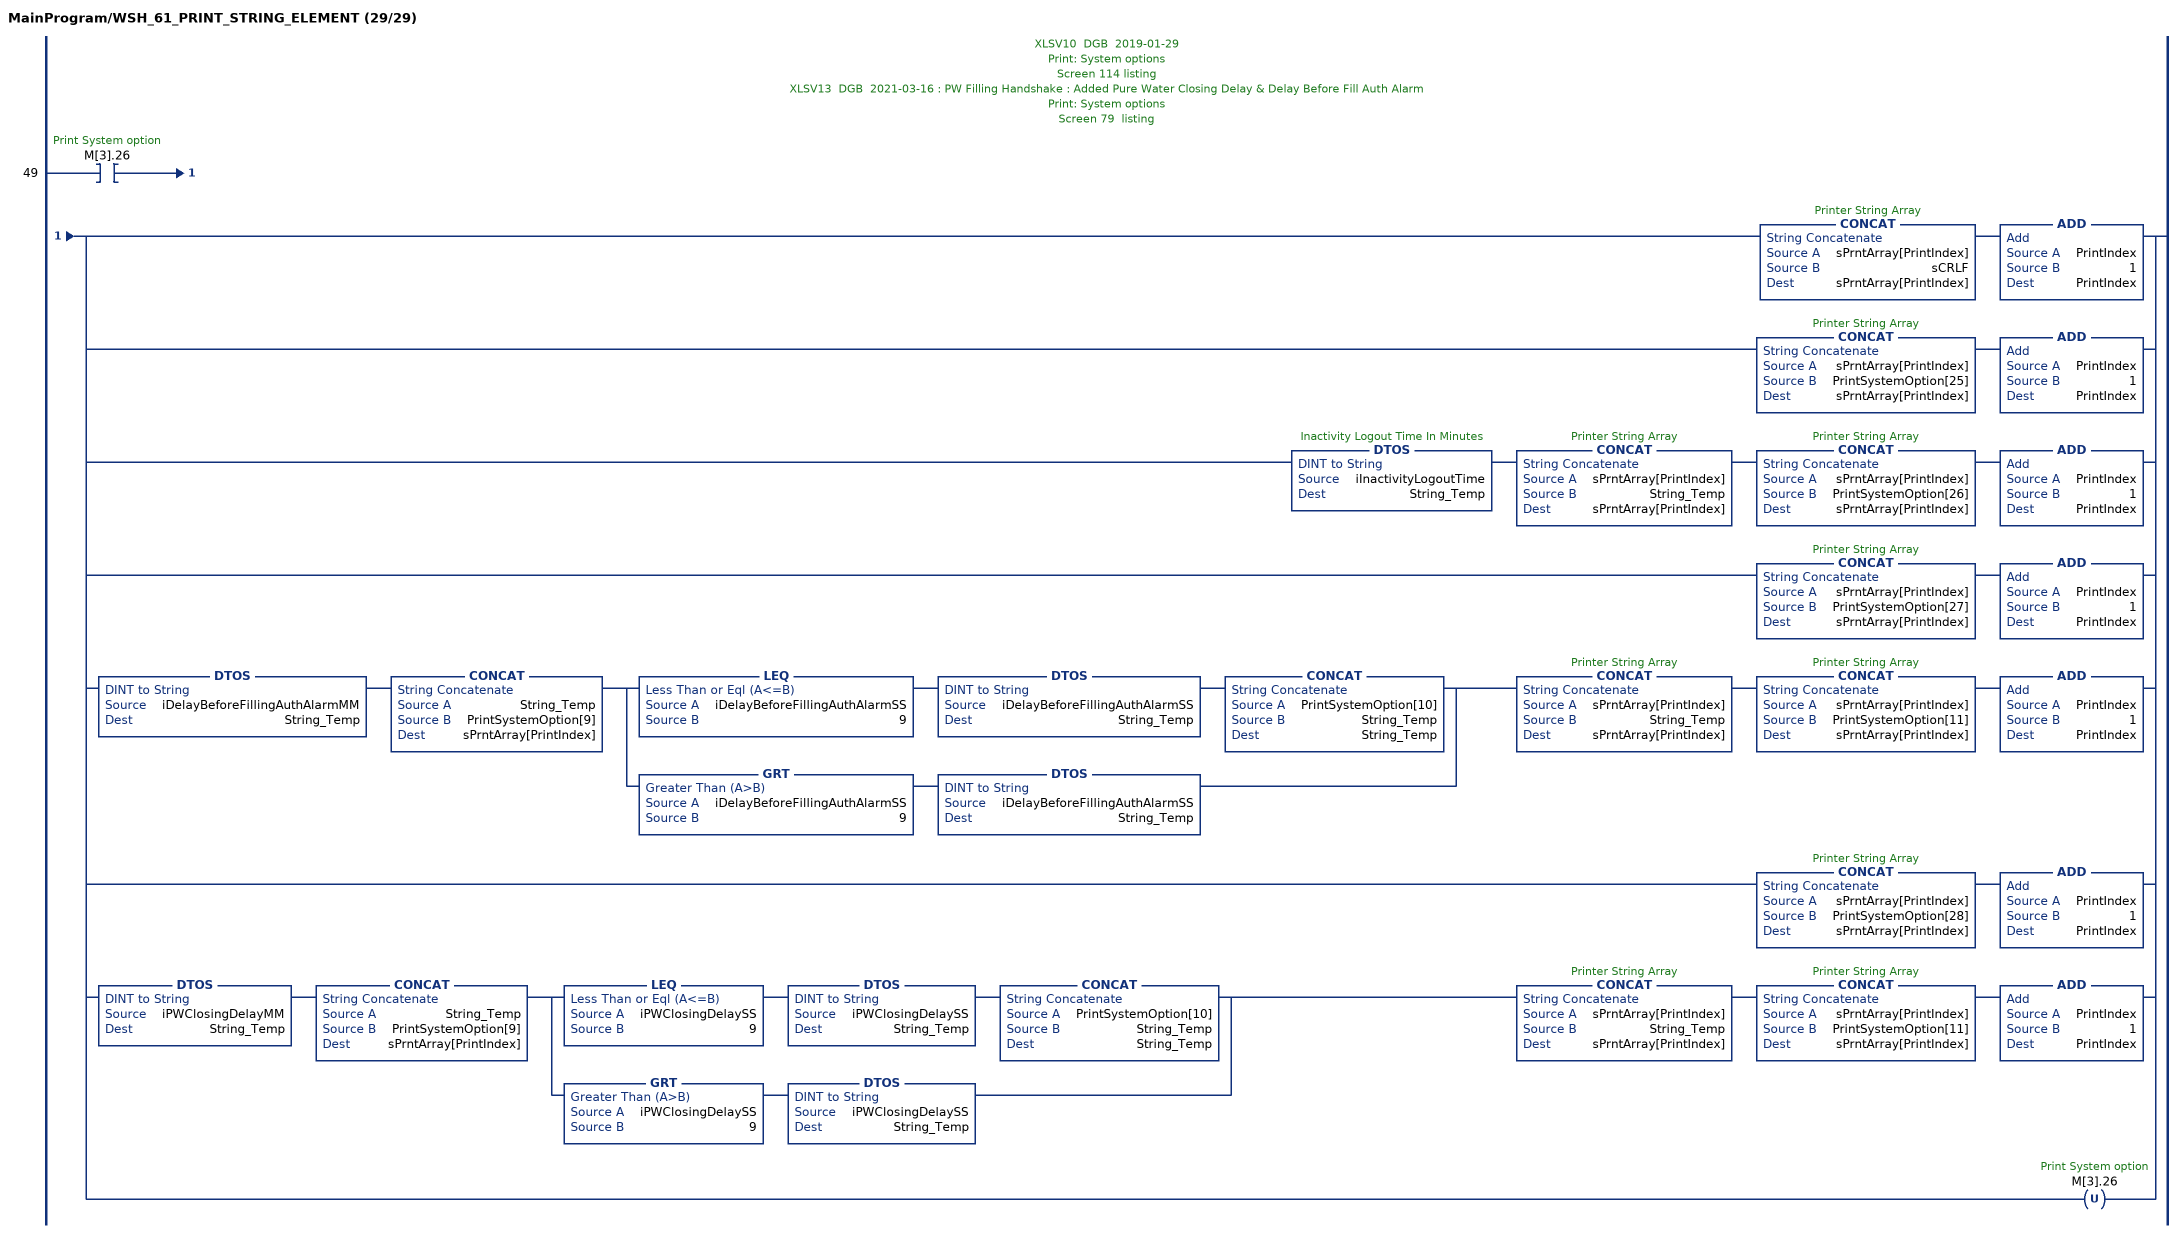
   // XLSV10  DGB  2019-01-29
   // Print: System options
   // Screen 114 listing
   // XLSV13  DGB  2021-03-16 : PW Filling Handshake : Added Pure Water Closing Delay & Delay Before Fill Auth Alarm
   // Print: System options
   // Screen 79  listing
   49: XIC(M[3].26)[CONCAT(sPrntArray[PrintIndex],sCRLF,sPrntArray[PrintIndex]) ADD(PrintIndex,1,PrintIndex) ,CONCAT(sPrntArray[PrintIndex],PrintSystemOption[25],sPrntArray[PrintIndex]) ADD(PrintIndex,1,PrintIndex) ,DTOS(iInactivityLogoutTime,String_Temp) CONCAT(sPrntArray[PrintIndex],String_Temp,sPrntArray[PrintIndex]) CONCAT(sPrntArray[PrintIndex],PrintSystemOption[26],sPrntArray[PrintIndex]) ADD(PrintIndex,1,PrintIndex) ,CONCAT(sPrntArray[PrintIndex],PrintSystemOption[27],sPrntArray[PrintIndex]) ADD(PrintIndex,1,PrintIndex) ,DTOS(iDelayBeforeFillingAuthAlarmMM,String_Temp) CONCAT(String_Temp,PrintSystemOption[9],sPrntArray[PrintIndex]) [LEQ(iDelayBeforeFillingAuthAlarmSS,9) DTOS(iDelayBeforeFillingAuthAlarmSS,String_Temp) CONCAT(PrintSystemOption[10],String_Temp,String_Temp) ,GRT(iDelayBeforeFillingAuthAlarmSS,9) DTOS(iDelayBeforeFillingAuthAlarmSS,String_Temp) ] CONCAT(sPrntArray[PrintIndex],String_Temp,sPrntArray[PrintIndex]) CONCAT(sPrntArray[PrintIndex],PrintSystemOption[11],sPrntArray[PrintIndex]) ADD(PrintIndex,1,PrintIndex) ,CONCAT(sPrntArray[PrintIndex],PrintSystemOption[28],sPrntArray[PrintIndex]) ADD(PrintIndex,1,PrintIndex) ,DTOS(iPWClosingDelayMM,String_Temp) CONCAT(String_Temp,PrintSystemOption[9],sPrntArray[PrintIndex]) [LEQ(iPWClosingDelaySS,9) DTOS(iPWClosingDelaySS,String_Temp) CONCAT(PrintSystemOption[10],String_Temp,String_Temp) ,GRT(iPWClosingDelaySS,9) DTOS(iPWClosingDelaySS,String_Temp) ] CONCAT(sPrntArray[PrintIndex],String_Temp,sPrntArray[PrintIndex]) CONCAT(sPrntArray[PrintIndex],PrintSystemOption[11],sPrntArray[PrintIndex]) ADD(PrintIndex,1,PrintIndex) ,OTU(M[3].26) ];
END_ROUTINE
